{region 'Documentation'}
(*!
<summary>Checks LREAL non-finite scalar operands and Error above held Failed.</summary>
<description>
Quiet NaN and both infinities are built by bit representation, never exceptional arithmetic.
Actual, expected/bound and tolerance roles are exercised separately across algorithm families.
NaNAfterFailure deliberately retains the preceding subject results; other rows reset them.
A disabled preparation call consumes subject resets before the next enabled observation.
Only outer checking Assertions contribute to the Test Case result.
Expected outcomes are explicit; production processing is inherited, not mirrored.
</description>
*)
{endregion}
FUNCTION_BLOCK Test_AssertionNonFinite_LReal EXTENDS TestCaseBase
VAR
    FEqualSubject : AssertEqual_LReal;
    FLessThanSubject : AssertLessThan_LReal;
    FInRangeSubject : AssertInRange_LReal;
    FEqualToleranceSubject : AssertEqualTolerance_LReal;
    FNotEqualToleranceSubject : AssertNotEqualTolerance_LReal;
    FActual : LREAL;
    FExpected : LREAL;
    FLower : LREAL;
    FUpper : LREAL;
    FTolerance : LREAL;
    FQuietNaN : FloatingPointBits_LReal;
    FPositiveInfinity : FloatingPointBits_LReal;
    FNegativeInfinity : FloatingPointBits_LReal;
    FExpectedEqualResult : E_Result;
    FExpectedLessThanResult : E_Result;
    FExpectedInRangeResult : E_Result;
    FExpectedEqualToleranceResult : E_Result;
    FExpectedNotEqualToleranceResult : E_Result;
    FExpectedFindings : UDINT;
    FCapture : EventBuffer;
    FEvents : ARRAY[1..CaptureLength] OF ST_Event;
    FCaptureFifo : ST_FifoStatus;
    FCaptureStatus : ST_EventBufferStatus;
    FRow : UINT;
    FRowPrepared : BOOL;
    FPreserveResults : BOOL;
    FObservationReady : BOOL;
    FChecked : BOOL;
    FSetupValid : BOOL;
END_VAR
VAR
    FEqualResult : AssertTrue;
    FEqualResultMatches : BOOL;
    FLessThanResult : AssertTrue;
    FLessThanResultMatches : BOOL;
    FInRangeResult : AssertTrue;
    FInRangeResultMatches : BOOL;
    FEqualToleranceResult : AssertTrue;
    FEqualToleranceResultMatches : BOOL;
    FNotEqualToleranceResult : AssertTrue;
    FNotEqualToleranceResultMatches : BOOL;
    FCaptureIntegrity : AssertTrue;
    FCaptureIntegrityMatches : BOOL;
    FFindingDetails : AssertTrue;
    FFindingDetailsMatch : BOOL;
END_VAR
VAR CONSTANT
    CaptureLength : UINT := 16;
    FixtureSize : UINT := 8;
    OneBits : LWORD := LWORD#16#3FF0000000000000;
    QuietNaNBits : LWORD := LWORD#16#7FF8000000000000;
    PositiveInfinityBits : LWORD := LWORD#16#7FF0000000000000;
    NegativeInfinityBits : LWORD := LWORD#16#FFF0000000000000;
    ActualQuietNaN : UINT := 1;
    ActualPositiveInfinity : UINT := 2;
    ActualNegativeInfinity : UINT := 3;
    ExpectedQuietNaN : UINT := 4;
    ExpectedPositiveInfinity : UINT := 5;
    ExpectedNegativeInfinity : UINT := 6;
    LowerBoundQuietNaN : UINT := 7;
    LowerBoundPositiveInfinity : UINT := 8;
    LowerBoundNegativeInfinity : UINT := 9;
    UpperBoundQuietNaN : UINT := 10;
    UpperBoundPositiveInfinity : UINT := 11;
    UpperBoundNegativeInfinity : UINT := 12;
    ToleranceQuietNaN : UINT := 13;
    TolerancePositiveInfinity : UINT := 14;
    ToleranceNegativeInfinity : UINT := 15;
    FailureBeforeNaN : UINT := 16;
    NaNAfterFailure : UINT := 17;
    LastRow : UINT := NaNAfterFailure;
END_VAR

SUPER^();

{region 'Documentation'}
(*!
<summary>Collects only outer checking Assertions, never intentional subject findings.</summary>
*)
{endregion}
METHOD PROTECTED AggregateResults
VAR_INPUT
    Aggregator : I_ResultAggregator; //! Borrowed result sink owned by the outer Test Case; add this test's checking Assertions without resetting or retaining the sink.
END_VAR
Aggregator.AddProvider(Provider := FEqualResult);
Aggregator.AddProvider(Provider := FLessThanResult);
Aggregator.AddProvider(Provider := FInRangeResult);
Aggregator.AddProvider(Provider := FEqualToleranceResult);
Aggregator.AddProvider(Provider := FNotEqualToleranceResult);
Aggregator.AddProvider(Provider := FCaptureIntegrity);
Aggregator.AddProvider(Provider := FFindingDetails);
END_METHOD

{region 'Documentation'}
(*!
<summary>Calls each inherited production Assertion once using the selected row.</summary>
*)
{endregion}
METHOD PRIVATE CallSubjects
VAR_INPUT
    Enable : BOOL; //! Observation-enable input forwarded to the controlled Assertion subjects for this call.
END_VAR
FEqualSubject(Enable := Enable,
    State := E_State.Running,
    IN := FActual,
    Expected := FExpected);
FLessThanSubject(Enable := Enable,
    State := E_State.Running,
    IN := FActual,
    Maximum := FExpected);
FInRangeSubject(Enable := Enable,
    State := E_State.Running,
    IN := FActual,
    Minimum := FLower,
    Maximum := FUpper);
FEqualToleranceSubject(Enable := Enable,
    State := E_State.Running,
    IN := FActual,
    Expected := FExpected,
    Tolerance := FTolerance);
FNotEqualToleranceSubject(Enable := Enable,
    State := E_State.Running,
    IN := FActual,
    Expected := FExpected,
    Tolerance := FTolerance);
END_METHOD

{region 'Documentation'}
(*!
<summary>Extends base validation with subject and checking-Assertion setup.</summary>
*)
{endregion}
METHOD PROTECTED CheckInitialization : BOOL //! TRUE when the inherited initialization check and this concrete fixture check both accept the setup.
CheckInitialization := SUPER^.CheckInitialization();
IF NOT CheckInitialization THEN
    RETURN;
END_IF;

CheckInitialization := FSetupValid
    AND FEqualResult.IsInitialized
    AND FLessThanResult.IsInitialized
    AND FInRangeResult.IsInitialized
    AND FEqualToleranceResult.IsInitialized
    AND FNotEqualToleranceResult.IsInitialized
    AND FCaptureIntegrity.IsInitialized
    AND FFindingDetails.IsInitialized;
IF NOT CheckInitialization THEN
    EventPublisher.PublishEvent(Event := CreateFrameworkEvent(Name := Name,
        ResourceName := '',
        State := State,
        Severity := E_EventSeverity.Error,
        Message := 'Floating-point selftest setup or fixture representation failed.'));
END_IF;
END_METHOD

{region 'Documentation'}
(*!
<summary>Checks literal results and the ordered isolated findings from this row.</summary>
*)
{endregion}
METHOD PRIVATE CheckResults
VAR
    FindingIndex : UINT;
    FindingMatches : BOOL;
END_VAR
FEqualResultMatches := FEqualSubject.Result = FExpectedEqualResult;
FLessThanResultMatches := FLessThanSubject.Result = FExpectedLessThanResult;
FInRangeResultMatches := FInRangeSubject.Result = FExpectedInRangeResult;
FEqualToleranceResultMatches := FEqualToleranceSubject.Result = FExpectedEqualToleranceResult;
FNotEqualToleranceResultMatches := FNotEqualToleranceSubject.Result = FExpectedNotEqualToleranceResult;
FCaptureIntegrityMatches := (FCaptureStatus.SequenceId = FExpectedFindings)
    AND (FCaptureStatus.LostEventCount = 0);

FindingIndex := 1;
FFindingDetailsMatch := TRUE;
IF (FExpectedEqualResult = E_Result.Failed) OR (FExpectedEqualResult = E_Result.Error) THEN
    FindingMatches := IsFindingValid(Index := FindingIndex,
        ExpectedName := FEqualSubject.Name,
        ExpectedResult := FExpectedEqualResult);
    FFindingDetailsMatch := FFindingDetailsMatch AND FindingMatches;
    FindingIndex := FindingIndex + 1;
END_IF;
IF (FExpectedLessThanResult = E_Result.Failed) OR (FExpectedLessThanResult = E_Result.Error) THEN
    FindingMatches := IsFindingValid(Index := FindingIndex,
        ExpectedName := FLessThanSubject.Name,
        ExpectedResult := FExpectedLessThanResult);
    FFindingDetailsMatch := FFindingDetailsMatch AND FindingMatches;
    FindingIndex := FindingIndex + 1;
END_IF;
IF (FExpectedInRangeResult = E_Result.Failed) OR (FExpectedInRangeResult = E_Result.Error) THEN
    FindingMatches := IsFindingValid(Index := FindingIndex,
        ExpectedName := FInRangeSubject.Name,
        ExpectedResult := FExpectedInRangeResult);
    FFindingDetailsMatch := FFindingDetailsMatch AND FindingMatches;
    FindingIndex := FindingIndex + 1;
END_IF;
IF (FExpectedEqualToleranceResult = E_Result.Failed) OR (FExpectedEqualToleranceResult = E_Result.Error) THEN
    FindingMatches := IsFindingValid(Index := FindingIndex,
        ExpectedName := FEqualToleranceSubject.Name,
        ExpectedResult := FExpectedEqualToleranceResult);
    FFindingDetailsMatch := FFindingDetailsMatch AND FindingMatches;
    FindingIndex := FindingIndex + 1;
END_IF;
IF (FExpectedNotEqualToleranceResult = E_Result.Failed) OR (FExpectedNotEqualToleranceResult = E_Result.Error) THEN
    FindingMatches := IsFindingValid(Index := FindingIndex,
        ExpectedName := FNotEqualToleranceSubject.Name,
        ExpectedResult := FExpectedNotEqualToleranceResult);
    FFindingDetailsMatch := FFindingDetailsMatch AND FindingMatches;
    FindingIndex := FindingIndex + 1;
END_IF;
END_METHOD

{region 'Documentation'}
(*!
<summary>Configures checking Assertions; subject actions remain in the test script.</summary>
*)
{endregion}
METHOD PROTECTED Configure
VAR
    Initialized : BOOL;
END_VAR
FPreparationStateCount := 0;
FTestStateCount := 1;
FSetupValid := InitializeValues();
FEqualResult.Initialize(Parent := THIS^,
    AssertionName := 'EqualResult');
FLessThanResult.Initialize(Parent := THIS^,
    AssertionName := 'LessThanResult');
FInRangeResult.Initialize(Parent := THIS^,
    AssertionName := 'InRangeResult');
FEqualToleranceResult.Initialize(Parent := THIS^,
    AssertionName := 'EqualToleranceResult');
FNotEqualToleranceResult.Initialize(Parent := THIS^,
    AssertionName := 'NotEqualToleranceResult');
FCaptureIntegrity.Initialize(Parent := THIS^,
    AssertionName := 'CaptureIntegrity');
FFindingDetails.Initialize(Parent := THIS^,
    AssertionName := 'FindingDetails');
Initialized := FCapture.Initialize(Buffer := FEvents,
    FifoControl := FCaptureFifo,
    Status := FCaptureStatus);
FSetupValid := FSetupValid AND Initialized;
FEqualSubject.BindPublisher(Publisher := FCapture);
Initialized := FEqualSubject.Initialize(Parent := THIS^,
    AssertionName := 'EqualSubject');
FSetupValid := FSetupValid AND Initialized;
FLessThanSubject.BindPublisher(Publisher := FCapture);
Initialized := FLessThanSubject.Initialize(Parent := THIS^,
    AssertionName := 'LessThanSubject');
FSetupValid := FSetupValid AND Initialized;
FInRangeSubject.BindPublisher(Publisher := FCapture);
Initialized := FInRangeSubject.Initialize(Parent := THIS^,
    AssertionName := 'InRangeSubject');
FSetupValid := FSetupValid AND Initialized;
FEqualToleranceSubject.BindPublisher(Publisher := FCapture);
Initialized := FEqualToleranceSubject.Initialize(Parent := THIS^,
    AssertionName := 'EqualToleranceSubject');
FSetupValid := FSetupValid AND Initialized;
FNotEqualToleranceSubject.BindPublisher(Publisher := FCapture);
Initialized := FNotEqualToleranceSubject.Initialize(Parent := THIS^,
    AssertionName := 'NotEqualToleranceSubject');
FSetupValid := FSetupValid AND Initialized;
END_METHOD

{region 'Documentation'}
(*!
<summary>Establishes typed fixtures and verifies their representation before any subject call.</summary>
*)
{endregion}
METHOD PRIVATE InitializeValues : BOOL //! TRUE when fixture sizes and floating-point bit representations match their explicit expected patterns.
VAR
    Representation : FloatingPointBits_LReal;
END_VAR
Representation.Value := LREAL#1.0;
InitializeValues := (SIZEOF(Representation) = FixtureSize)
    AND (Representation.Bits = OneBits);

FQuietNaN.Bits := QuietNaNBits;
Representation.Value := FQuietNaN.Value;
InitializeValues := InitializeValues AND (Representation.Bits = QuietNaNBits);
FPositiveInfinity.Bits := PositiveInfinityBits;
Representation.Value := FPositiveInfinity.Value;
InitializeValues := InitializeValues AND (Representation.Bits = PositiveInfinityBits);
FNegativeInfinity.Bits := NegativeInfinityBits;
Representation.Value := FNegativeInfinity.Value;
InitializeValues := InitializeValues AND (Representation.Bits = NegativeInfinityBits);
END_METHOD

{region 'Documentation'}
(*!
<summary>Reads a captured finding; the caller bounds the index by 5 subjects.</summary>
*)
{endregion}
METHOD PRIVATE IsFindingValid : BOOL //! TRUE when the selected captured finding satisfies the scenario metadata and diagnostic checks.
VAR_INPUT
    Index : UINT; //! One-based index in the retained isolated event capture.
    ExpectedName : STRING(GVL_Constants.NameLength); //! Independently authored Assertion name expected in the selected finding.
    ExpectedResult : E_Result; //! Independently authored finding result.
END_VAR
IsFindingValid := (FEvents[Index].SequenceId = UINT_TO_UDINT(Index))
    AND (FEvents[Index].Name = ExpectedName)
    AND (FEvents[Index].OwnerScope = E_OwnerScope.Assertion)
    AND (FEvents[Index].EventType = E_EventType.Result)
    AND (FEvents[Index].State = E_State.Running)
    AND (FEvents[Index].Result = ExpectedResult)
    AND (FEvents[Index].Message <> '');
END_METHOD

{region 'Documentation'}
(*!
<summary>Completes abort without asynchronous resources.</summary>
*)
{endregion}
METHOD PROTECTED ProcessAbort
VAR_INPUT
    Enable : BOOL; //! Phase permission supplied by the owning Test Case; FALSE does not authorize progression, while observation may continue.
END_VAR
IF Enable THEN
    CompleteAbort();
END_IF;
END_METHOD

{region 'Documentation'}
(*!
<summary>Latches checked observations before the next script step may proceed.</summary>
*)
{endregion}
METHOD PROTECTED ProcessAssertions
VAR_INPUT
    Enable : BOOL; //! Phase permission supplied by the owning Test Case; FALSE does not authorize progression, while observation may continue.
END_VAR
VAR
    Evaluate : BOOL;
END_VAR
Evaluate := Enable AND FObservationReady;
FEqualResult(Enable := Evaluate,
    State := State,
    IN := FEqualResultMatches);
FLessThanResult(Enable := Evaluate,
    State := State,
    IN := FLessThanResultMatches);
FInRangeResult(Enable := Evaluate,
    State := State,
    IN := FInRangeResultMatches);
FEqualToleranceResult(Enable := Evaluate,
    State := State,
    IN := FEqualToleranceResultMatches);
FNotEqualToleranceResult(Enable := Evaluate,
    State := State,
    IN := FNotEqualToleranceResultMatches);
FCaptureIntegrity(Enable := Evaluate,
    State := State,
    IN := FCaptureIntegrityMatches);
FFindingDetails(Enable := Evaluate,
    State := State,
    IN := FFindingDetailsMatch);
IF Evaluate THEN
    FChecked := TRUE;
END_IF;
END_METHOD

{region 'Documentation'}
(*!
<summary>No Preparation phase is required.</summary>
*)
{endregion}
METHOD PROTECTED ProcessPreparations
VAR_INPUT
    // SA0033: Required hook; this test has no Preparation phase.
    {attribute 'analysis' := '-33'}
    Enable : BOOL; //! Phase permission supplied by the owning Test Case; FALSE does not authorize progression, while observation may continue.
END_VAR
END_METHOD

{region 'Documentation'}
(*!
<summary>Restarts the script and resets the checking Assertions.</summary>
*)
{endregion}
METHOD PROTECTED ProcessReset
FRow := ActualQuietNaN;
FRowPrepared := FALSE;
FChecked := FALSE;
FObservationReady := FALSE;
FEqualResult.Reset();
FEqualResultMatches := TRUE;
FLessThanResult.Reset();
FLessThanResultMatches := TRUE;
FInRangeResult.Reset();
FInRangeResultMatches := TRUE;
FEqualToleranceResult.Reset();
FEqualToleranceResultMatches := TRUE;
FNotEqualToleranceResult.Reset();
FNotEqualToleranceResultMatches := TRUE;
FCaptureIntegrity.Reset();
FCaptureIntegrityMatches := TRUE;
FFindingDetails.Reset();
FFindingDetailsMatch := TRUE;
CompleteReset();
END_METHOD

{region 'Documentation'}
(*!
<summary>Advances one bounded script step per active PLC cycle.</summary>
*)
{endregion}
METHOD PROTECTED ProcessTests
VAR_INPUT
    Enable : BOOL; //! Phase permission supplied by the owning Test Case; FALSE does not authorize progression, while observation may continue.
END_VAR
IF NOT Enable THEN
    RETURN;
END_IF;

IF FChecked THEN
    FChecked := FALSE;
    FObservationReady := FALSE;
    IF FRow = LastRow THEN
        CompleteTests();
        RETURN;
    END_IF;
    FRow := FRow + 1;
    FRowPrepared := FALSE;
END_IF;

IF NOT FRowPrepared THEN
    SelectRow();
    FCapture.Reset();
    IF NOT FPreserveResults THEN
        ResetSubjects();
    END_IF;
    CallSubjects(Enable := FALSE);
    FRowPrepared := TRUE;
ELSE
    CallSubjects(Enable := TRUE);
    CheckResults();
    FObservationReady := TRUE;
END_IF;
END_METHOD

{region 'Documentation'}
(*!
<summary>Requests fresh subject results before the next disabled call.</summary>
*)
{endregion}
METHOD PRIVATE ResetSubjects
FEqualSubject.Reset();
FLessThanSubject.Reset();
FInRangeSubject.Reset();
FEqualToleranceSubject.Reset();
FNotEqualToleranceSubject.Reset();
END_METHOD

{region 'Documentation'}
(*!
<summary>Selects independent literal outcomes; only named escalation rows preserve results.</summary>
*)
{endregion}
METHOD PRIVATE SelectRow
FPreserveResults := FALSE;
CASE FRow OF
    ActualQuietNaN:
        FActual := FQuietNaN.Value;
        FExpected := LREAL#1.0;
        FLower := LREAL#0.0;
        FUpper := LREAL#2.0;
        FTolerance := LREAL#0.5;
        FExpectedEqualResult := E_Result.Error;
        FExpectedLessThanResult := E_Result.Error;
        FExpectedInRangeResult := E_Result.Error;
        FExpectedEqualToleranceResult := E_Result.Error;
        FExpectedNotEqualToleranceResult := E_Result.Error;
        FExpectedFindings := 5;
    ActualPositiveInfinity:
        FActual := FPositiveInfinity.Value;
        FExpected := LREAL#1.0;
        FLower := LREAL#0.0;
        FUpper := LREAL#2.0;
        FTolerance := LREAL#0.5;
        FExpectedEqualResult := E_Result.Error;
        FExpectedLessThanResult := E_Result.Error;
        FExpectedInRangeResult := E_Result.Error;
        FExpectedEqualToleranceResult := E_Result.Error;
        FExpectedNotEqualToleranceResult := E_Result.Error;
        FExpectedFindings := 5;
    ActualNegativeInfinity:
        FActual := FNegativeInfinity.Value;
        FExpected := LREAL#1.0;
        FLower := LREAL#0.0;
        FUpper := LREAL#2.0;
        FTolerance := LREAL#0.5;
        FExpectedEqualResult := E_Result.Error;
        FExpectedLessThanResult := E_Result.Error;
        FExpectedInRangeResult := E_Result.Error;
        FExpectedEqualToleranceResult := E_Result.Error;
        FExpectedNotEqualToleranceResult := E_Result.Error;
        FExpectedFindings := 5;
    ExpectedQuietNaN:
        FActual := LREAL#1.0;
        FExpected := FQuietNaN.Value;
        FLower := LREAL#0.0;
        FUpper := LREAL#2.0;
        FTolerance := LREAL#0.5;
        FExpectedEqualResult := E_Result.Error;
        FExpectedLessThanResult := E_Result.Error;
        FExpectedInRangeResult := E_Result.Passed;
        FExpectedEqualToleranceResult := E_Result.Error;
        FExpectedNotEqualToleranceResult := E_Result.Error;
        FExpectedFindings := 4;
    ExpectedPositiveInfinity:
        FActual := LREAL#1.0;
        FExpected := FPositiveInfinity.Value;
        FLower := LREAL#0.0;
        FUpper := LREAL#2.0;
        FTolerance := LREAL#0.5;
        FExpectedEqualResult := E_Result.Error;
        FExpectedLessThanResult := E_Result.Error;
        FExpectedInRangeResult := E_Result.Passed;
        FExpectedEqualToleranceResult := E_Result.Error;
        FExpectedNotEqualToleranceResult := E_Result.Error;
        FExpectedFindings := 4;
    ExpectedNegativeInfinity:
        FActual := LREAL#1.0;
        FExpected := FNegativeInfinity.Value;
        FLower := LREAL#0.0;
        FUpper := LREAL#2.0;
        FTolerance := LREAL#0.5;
        FExpectedEqualResult := E_Result.Error;
        FExpectedLessThanResult := E_Result.Error;
        FExpectedInRangeResult := E_Result.Passed;
        FExpectedEqualToleranceResult := E_Result.Error;
        FExpectedNotEqualToleranceResult := E_Result.Error;
        FExpectedFindings := 4;
    LowerBoundQuietNaN:
        FActual := LREAL#1.0;
        FExpected := LREAL#1.0;
        FLower := FQuietNaN.Value;
        FUpper := LREAL#2.0;
        FTolerance := LREAL#0.5;
        FExpectedEqualResult := E_Result.Passed;
        FExpectedLessThanResult := E_Result.Failed;
        FExpectedInRangeResult := E_Result.Error;
        FExpectedEqualToleranceResult := E_Result.Passed;
        FExpectedNotEqualToleranceResult := E_Result.Failed;
        FExpectedFindings := 3;
    LowerBoundPositiveInfinity:
        FActual := LREAL#1.0;
        FExpected := LREAL#1.0;
        FLower := FPositiveInfinity.Value;
        FUpper := LREAL#2.0;
        FTolerance := LREAL#0.5;
        FExpectedEqualResult := E_Result.Passed;
        FExpectedLessThanResult := E_Result.Failed;
        FExpectedInRangeResult := E_Result.Error;
        FExpectedEqualToleranceResult := E_Result.Passed;
        FExpectedNotEqualToleranceResult := E_Result.Failed;
        FExpectedFindings := 3;
    LowerBoundNegativeInfinity:
        FActual := LREAL#1.0;
        FExpected := LREAL#1.0;
        FLower := FNegativeInfinity.Value;
        FUpper := LREAL#2.0;
        FTolerance := LREAL#0.5;
        FExpectedEqualResult := E_Result.Passed;
        FExpectedLessThanResult := E_Result.Failed;
        FExpectedInRangeResult := E_Result.Error;
        FExpectedEqualToleranceResult := E_Result.Passed;
        FExpectedNotEqualToleranceResult := E_Result.Failed;
        FExpectedFindings := 3;
    UpperBoundQuietNaN:
        FActual := LREAL#1.0;
        FExpected := LREAL#1.0;
        FLower := LREAL#0.0;
        FUpper := FQuietNaN.Value;
        FTolerance := LREAL#0.5;
        FExpectedEqualResult := E_Result.Passed;
        FExpectedLessThanResult := E_Result.Failed;
        FExpectedInRangeResult := E_Result.Error;
        FExpectedEqualToleranceResult := E_Result.Passed;
        FExpectedNotEqualToleranceResult := E_Result.Failed;
        FExpectedFindings := 3;
    UpperBoundPositiveInfinity:
        FActual := LREAL#1.0;
        FExpected := LREAL#1.0;
        FLower := LREAL#0.0;
        FUpper := FPositiveInfinity.Value;
        FTolerance := LREAL#0.5;
        FExpectedEqualResult := E_Result.Passed;
        FExpectedLessThanResult := E_Result.Failed;
        FExpectedInRangeResult := E_Result.Error;
        FExpectedEqualToleranceResult := E_Result.Passed;
        FExpectedNotEqualToleranceResult := E_Result.Failed;
        FExpectedFindings := 3;
    UpperBoundNegativeInfinity:
        FActual := LREAL#1.0;
        FExpected := LREAL#1.0;
        FLower := LREAL#0.0;
        FUpper := FNegativeInfinity.Value;
        FTolerance := LREAL#0.5;
        FExpectedEqualResult := E_Result.Passed;
        FExpectedLessThanResult := E_Result.Failed;
        FExpectedInRangeResult := E_Result.Error;
        FExpectedEqualToleranceResult := E_Result.Passed;
        FExpectedNotEqualToleranceResult := E_Result.Failed;
        FExpectedFindings := 3;
    ToleranceQuietNaN:
        FActual := LREAL#1.0;
        FExpected := LREAL#1.0;
        FLower := LREAL#0.0;
        FUpper := LREAL#2.0;
        FTolerance := FQuietNaN.Value;
        FExpectedEqualResult := E_Result.Passed;
        FExpectedLessThanResult := E_Result.Failed;
        FExpectedInRangeResult := E_Result.Passed;
        FExpectedEqualToleranceResult := E_Result.Error;
        FExpectedNotEqualToleranceResult := E_Result.Error;
        FExpectedFindings := 3;
    TolerancePositiveInfinity:
        FActual := LREAL#1.0;
        FExpected := LREAL#1.0;
        FLower := LREAL#0.0;
        FUpper := LREAL#2.0;
        FTolerance := FPositiveInfinity.Value;
        FExpectedEqualResult := E_Result.Passed;
        FExpectedLessThanResult := E_Result.Failed;
        FExpectedInRangeResult := E_Result.Passed;
        FExpectedEqualToleranceResult := E_Result.Error;
        FExpectedNotEqualToleranceResult := E_Result.Error;
        FExpectedFindings := 3;
    ToleranceNegativeInfinity:
        FActual := LREAL#1.0;
        FExpected := LREAL#1.0;
        FLower := LREAL#0.0;
        FUpper := LREAL#2.0;
        FTolerance := FNegativeInfinity.Value;
        FExpectedEqualResult := E_Result.Passed;
        FExpectedLessThanResult := E_Result.Failed;
        FExpectedInRangeResult := E_Result.Passed;
        FExpectedEqualToleranceResult := E_Result.Error;
        FExpectedNotEqualToleranceResult := E_Result.Error;
        FExpectedFindings := 3;
    FailureBeforeNaN:
        FActual := LREAL#3.0;
        FExpected := LREAL#1.0;
        FLower := LREAL#0.0;
        FUpper := LREAL#2.0;
        FTolerance := LREAL#0.5;
        FExpectedEqualResult := E_Result.Failed;
        FExpectedLessThanResult := E_Result.Failed;
        FExpectedInRangeResult := E_Result.Failed;
        FExpectedEqualToleranceResult := E_Result.Failed;
        FExpectedNotEqualToleranceResult := E_Result.Passed;
        FExpectedFindings := 4;
    NaNAfterFailure:
        FActual := FQuietNaN.Value;
        FExpected := LREAL#1.0;
        FLower := LREAL#0.0;
        FUpper := LREAL#2.0;
        FTolerance := LREAL#0.5;
        FExpectedEqualResult := E_Result.Error;
        FExpectedLessThanResult := E_Result.Error;
        FExpectedInRangeResult := E_Result.Error;
        FExpectedEqualToleranceResult := E_Result.Error;
        FExpectedNotEqualToleranceResult := E_Result.Error;
        FExpectedFindings := 5;
        FPreserveResults := TRUE;
ELSE
    Error(Message := 'Unknown floating-point test row.');
END_CASE;
END_METHOD

END_FUNCTION_BLOCK

(* stored: Version 1.1.0.1
   POU Test_AssertionNonFinite_LReal: Id {5501ccff-29ae-495b-8c12-0543e82b3d63}, SpecialFunc None
   Folder Internal: Id {621f2a90-d955-4b4b-b80e-7d5b20138472}
   Method AggregateResults: Id {dcfd30a6-f91e-4743-8175-31ddc41a2f49}
   Method CallSubjects: Id {17585cdc-fb84-4494-b46c-70a4bf20832c}
   Method CheckInitialization: Id {eb8e31ed-2bf0-4fc6-866a-a9759b21c5dd}
   Method CheckResults: Id {b5f25e7b-4c13-4701-9d1f-4b7bafb7fa3f}
   Method Configure: Id {e2848a75-8a9a-40a9-8ca9-b3fe7b2fd4e6}
   Method InitializeValues: Id {81d70017-3e81-4132-9871-e14d505fdefa}
   Method IsFindingValid: Id {9afd6e1b-04e3-44b7-97c3-423f0f028c25}
   Method ProcessAbort: Id {088b5f26-5f0c-4abd-b7c6-cfa861a43d19}
   Method ProcessAssertions: Id {49e83692-b8a9-455c-bb86-13de344bfeb3}
   Method ProcessPreparations: Id {710fdb2e-ade5-454d-b77e-4dfe96b81046}
   Method ProcessReset: Id {621df69e-b202-4d41-aad7-1afb8bf2c396}
   Method ProcessTests: Id {68dfa479-30bb-4d2e-8406-7af271922458}
   Method ResetSubjects: Id {6ae7047e-9772-4d8f-be45-7baa36a1fbe1}
   Method SelectRow: Id {6eb885de-17da-424b-81dc-738fdb0d90b4} *)
